TYPE ST_PolarIIChamber_CupServiceCtrl :
STRUCT
	Lift : ST_PolarIIChamber_CupLiftServiceCtrl;
	Drainer : ST_PolarIIChamber_SelectThreeServiceCtrl;
END_STRUCT
END_TYPE

(* stored: Version 1.1.0.1, ProductVersion 3.1.4026.18
   DUT ST_PolarIIChamber_CupServiceCtrl: Id {14000000-0000-0000-0000-000000000061} *)
